PROGRAM Main
VAR
	fbFastBlinkTimerOff  : TON;
    fbFastBlinkTimerOn   : TON;
    tFastBlinkOffTime    : TIME := T#1000MS; // Mappable off-time
    tFastBlinkOnTime     : TIME := T#1000MS; // Mappable on-time
    bFastBlinkOn  : BOOL;
	bFastBlinkOff : BOOL;
	bFault : BOOL;
	bfault_EstopDiscrepancy : BOOL;
	bfault_FaultResetNCDiscrepancy : BOOL;
	bfault_FaultResetNODiscrepancy : BOOL;
	tDiscrepancyTimer : TIME := T#500MS;
	fbFaultRstNCDiscrepancyTimer: TON;
	fbFaultRstNODiscrepancyTimer: TON;
END_VAR

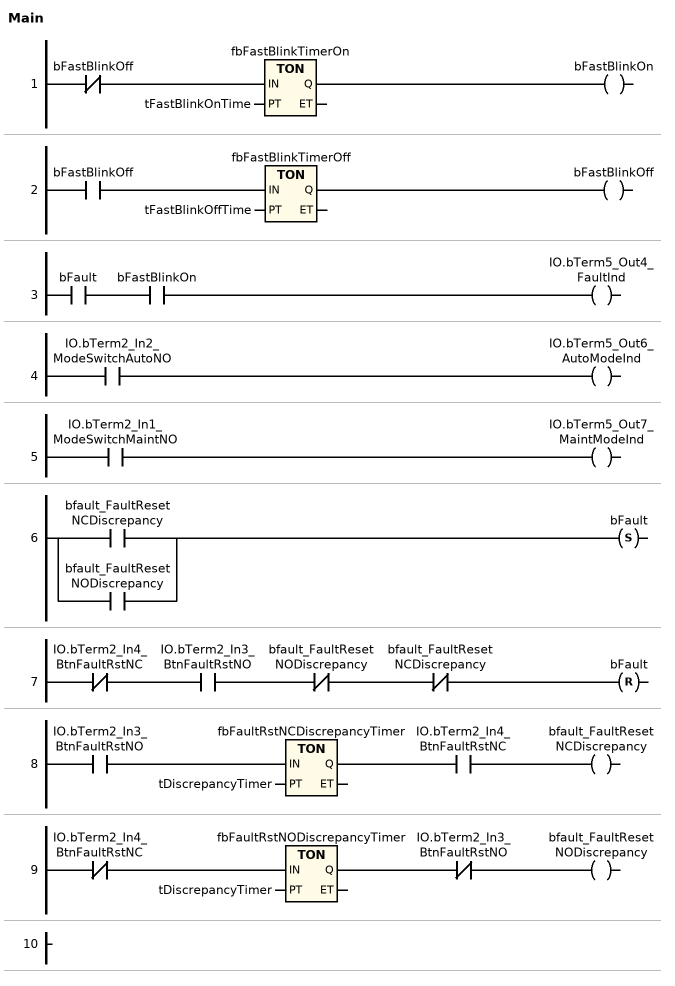
// NETWORK 1
fbFastBlinkTimerOn(IN := NOT bFastBlinkOff, PT := tFastBlinkOnTime); // TON
bFastBlinkOn := fbFastBlinkTimerOn.Q;

// NETWORK 2
fbFastBlinkTimerOff(IN := bFastBlinkOff, PT := tFastBlinkOffTime); // TON
bFastBlinkOff := fbFastBlinkTimerOff.Q;

// NETWORK 3
IO.bTerm5_Out4_FaultInd := bFault AND bFastBlinkOn;

// NETWORK 4
IO.bTerm5_Out6_AutoModeInd := IO.bTerm2_In2_ModeSwitchAutoNO;

// NETWORK 5
IO.bTerm5_Out7_MaintModeInd := IO.bTerm2_In1_ModeSwitchMaintNO;

// NETWORK 6
bFault S= bfault_FaultResetNCDiscrepancy OR bfault_FaultResetNODiscrepancy;

// NETWORK 7
bFault R= NOT IO.bTerm2_In4_BtnFaultRstNC AND IO.bTerm2_In3_BtnFaultRstNO AND NOT bfault_FaultResetNODiscrepancy AND NOT bfault_FaultResetNCDiscrepancy;

// NETWORK 8
fbFaultRstNCDiscrepancyTimer(IN := IO.bTerm2_In3_BtnFaultRstNO, PT := tDiscrepancyTimer); // TON
bfault_FaultResetNCDiscrepancy := fbFaultRstNCDiscrepancyTimer.Q AND IO.bTerm2_In4_BtnFaultRstNC;

// NETWORK 9
fbFaultRstNODiscrepancyTimer(IN := NOT IO.bTerm2_In4_BtnFaultRstNC, PT := tDiscrepancyTimer); // TON
bfault_FaultResetNODiscrepancy := fbFaultRstNODiscrepancyTimer.Q AND NOT IO.bTerm2_In3_BtnFaultRstNO;

// NETWORK 10

END_PROGRAM

(* stored: Version 1.1.0.1, ProductVersion 3.1.4024.16
   POU Main: Id {7cf0928f-9d39-4b48-8542-e2949f969e22}, SpecialFunc None *)
